Exceptions.ThrowGenericConversionNotSupported(
	sourceNamespaceName := NamespaceName,
	sourceClassName := ClassName,
	sourcePOUName := __POUNAME(),
	sourcePosition := __POSITION(),
	sourceDataType := TypeClass,
	targetDataType := otherValue.TypeClass
);
END_METHOD

(*!
<summary>Copies the stored byte representation into an equally sized target.</summary>
<description>
Requires a live writable target whose size equals Size. The caller is responsible for data compatibility: no
type check or numeric conversion is performed. Copies bytes from a nonzero Address referencing live source
storage. Does not clone referenced objects, transfer ownership, retain the target or modify this descriptor.
Copied pointer values still refer to the same resources and do not grant an independent right to release them.
A zero source Address raises DataMemberNotSpecifiedException without changing the target. A null target raises
ArgumentNotSpecifiedException; a target smaller than Size raises TargetVariableMemoryOverflowException; a
target larger than Size raises ArgumentOutOfRangeException before copying. Overlapping source and target
regions, including identical addresses, are supported through MEMMOVE. Descendants cannot override this
descriptor operation; customize value equality through IEqualityComparer or the stored object equality
contract.
</description>
*)
//!<param name="target">
//! Writable destination with the same byte size; its type interpretation is the caller's responsibility.
//! </param>
METHOD FINAL CopyTo
VAR_INPUT
	target : ANY;
END_VAR
IF Address = 0 THEN
	Exceptions.ThrowDataMemberNotSpecified(
		sourceNamespaceName := NamespaceName,
		sourceClassName := ClassName,
		sourcePOUName := __POUNAME(),
		sourcePosition := __POSITION(),
		dataMemberName := 'Address'
	);
END_IF

IF target.pValue = 0 THEN
	Exceptions.ThrowArgumentNotSpecified(
		sourceNamespaceName := NamespaceName,
		sourceClassName := ClassName,
		sourcePOUName := __POUNAME(),
		sourcePosition := __POSITION(),
		argumentName := 'target'
	); 
END_IF

IF TO_ULINT(target.diSize) < Size THEN
	Exceptions.ThrowTargetVariableMemoryOverflow(
		sourceNamespaceName := NamespaceName,
		sourceClassName := ClassName,
		sourcePOUName := __POUNAME(),
		sourcePosition := __POSITION(),
		targetVariableName := 'target.diSize',
		targetVariableSize := TO_ULINT(target.diSize)
	);
ELSIF TO_ULINT(target.diSize) > Size THEN
	Exceptions.ThrowArgumentOutOfRange(
		sourceNamespaceName := NamespaceName,
		sourceClassName := ClassName,
		sourcePOUName := __POUNAME(),
		sourcePosition := __POSITION(),
		argumentName := 'target.diSize',
		argumentValue := target.diSize
	);
END_IF

internalCopyTo(targetAddress := target.pValue);
END_METHOD

(*!
<summary>Compares generic values using an optional comparer or the built-in equality rules.</summary>
<description>
When comparer is supplied, AreEqual receives copies of both GENERIC_VALUE descriptors before any built-in
empty or type checks. OBJECT and USER_DEFINED remain distinct and Size is passed without conversion to
AnyType. The caller selects a compatible equality strategy, including its treatment of empty operands, and
keeps it and the data alive for the call. Comparer exceptions propagate without fallback. The comparer and
operands are borrowed only for the call; no payload is copied, cloned or released, and no ownership is
transferred. IsMemoryOwner does not affect the strategy's equality result. A supplied strategy must provide
GetValueHashCode consistent with AreEqual; this method does not compute a hash. Without a comparer, the
following built-in rules apply. INT_8 through INT_64 and UINT_8 through UINT_64 compare by value across widths
and signedness without floating-point conversion. A negative signed value never equals an unsigned value.
Pairs of REAL_32/REAL_64 values compare by canonical binary64 representation after widening non-NaN REAL
values, without a tolerance: positive and negative zero are equal, and all NaN encodings compare equal to each
other, including across widths, but not to non-NaN values. NaN is classified from integer bit views before
widening; other REAL widening follows the runtime floating-point configuration. A nonempty integer value and a
nonempty floating-point value always compare unequal, in either operand order. Both empty descriptors compare
equal; one empty descriptor compares unequal to a nonempty one. For nonempty descriptors, different TypeClass
values compare unequal except for the integer and floating-point pairs described above. BOOLEAN values compare
logically. Nonempty OBJECT descriptors delegate to the first live Object instance's Equals with the second
instance as its argument. The object type must provide a symmetric, transitive equality relation and a
matching GetHashCode; base Object uses identity equality. Callbacks and their exceptions propagate without
fallback. An address does not validate object lifetime. Other matching categories retain byte comparison:
strings use their actual string sizes, otherwise descriptor sizes are used. Dates and times compare by
representation only within the same TypeClass. Byte comparison covers the full ULINT length in bounded MEMCMP
chunks. USER_DEFINED compares all Size bytes, including padding and stored pointer values; equal fields do not
necessarily imply equal bytes, and the concrete user-defined type identity is not checked. Supply a compatible
comparer for field-based equality. Both descriptors must reference live storage consistent with their type and
size; no ownership is transferred. Descendants cannot override this descriptor operation; customize value
equality through IEqualityComparer or the stored object equality contract.
</description>
*)
//!<param name="otherValue">Descriptor of the value to compare.</param>
//!<param name="comparer">Optional borrowed equality and hashing strategy; zero selects built-in equality.</param>
METHOD FINAL Equals : BOOL
VAR_INPUT
	otherValue : GENERIC_VALUE;
	comparer : IEqualityComparer := 0;
END_VAR
VAR
	signedValue : LINT;

	firstObject : POINTER TO Object;
	secondObject : POINTER TO Object;

	stringPointer : POINTER TO STRING;
	wideStringPointer : POINTER TO WSTRING;
	referenceDataSize : ULINT;
	valueToCompareDataSize : ULINT;
	comparedSize : ULINT;
	chunkSize : UDINT;
END_VAR
IF comparer <> 0 THEN
	Equals := comparer.AreEqual(first := THIS^, second := otherValue);
	
	RETURN;
END_IF

IF IsNull OR_ELSE otherValue.IsNull THEN
	Equals := IsNull AND_THEN otherValue.IsNull;
ELSE
	CASE TypeClass OF
		GENERIC_TYPE_CLASS.INT_8, GENERIC_TYPE_CLASS.INT_16, GENERIC_TYPE_CLASS.INT_32, GENERIC_TYPE_CLASS.INT_64:
			CASE otherValue.TypeClass OF
				GENERIC_TYPE_CLASS.INT_8, GENERIC_TYPE_CLASS.INT_16, GENERIC_TYPE_CLASS.INT_32, GENERIC_TYPE_CLASS.INT_64:
					Equals := AsLInt() = otherValue.AsLInt();
					RETURN;

				GENERIC_TYPE_CLASS.UINT_8, GENERIC_TYPE_CLASS.UINT_16, GENERIC_TYPE_CLASS.UINT_32, GENERIC_TYPE_CLASS.UINT_64:
					signedValue := AsLInt();
					Equals := signedValue >= SignedInt64.ZERO AND_THEN TO_ULINT(signedValue) = otherValue.AsULInt();
					RETURN;
			END_CASE

		GENERIC_TYPE_CLASS.UINT_8, GENERIC_TYPE_CLASS.UINT_16, GENERIC_TYPE_CLASS.UINT_32, GENERIC_TYPE_CLASS.UINT_64:
			CASE otherValue.TypeClass OF
				GENERIC_TYPE_CLASS.INT_8, GENERIC_TYPE_CLASS.INT_16, GENERIC_TYPE_CLASS.INT_32, GENERIC_TYPE_CLASS.INT_64:
					signedValue := otherValue.AsLInt();
					Equals := signedValue >= SignedInt64.ZERO AND_THEN AsULInt() = TO_ULINT(signedValue);
					RETURN;

				GENERIC_TYPE_CLASS.UINT_8, GENERIC_TYPE_CLASS.UINT_16, GENERIC_TYPE_CLASS.UINT_32, GENERIC_TYPE_CLASS.UINT_64:
					Equals := AsULInt() = otherValue.AsULInt();
					RETURN;
			END_CASE

		GENERIC_TYPE_CLASS.REAL_32, GENERIC_TYPE_CLASS.REAL_64:
			CASE otherValue.TypeClass OF
				GENERIC_TYPE_CLASS.REAL_32, GENERIC_TYPE_CLASS.REAL_64:
					Equals := getCanonicalRealBits() = otherValue.getCanonicalRealBits();
					RETURN;
			END_CASE
	END_CASE

	IF TypeClass <> otherValue.TypeClass THEN
		Equals := FALSE;
		RETURN;
	END_IF

	IF TypeClass = GENERIC_TYPE_CLASS.OBJECT THEN
		firstObject := Address;
		secondObject := otherValue.Address;
		Equals := firstObject^.Equals(other := secondObject^);
		RETURN;
	END_IF

	IF TypeClass = GENERIC_TYPE_CLASS.BOOLEAN THEN
		Equals := AsBool() = otherValue.AsBool();
		RETURN;
	END_IF

	IF TypeClass = GENERIC_TYPE_CLASS.STRING_8 AND_THEN otherValue.TypeClass = GENERIC_TYPE_CLASS.STRING_8 THEN
		stringPointer := Address;
		referenceDataSize := Strings.GetActualSize(value := stringPointer^);
		
		stringPointer := otherValue.Address;		
		valueToCompareDataSize := Strings.GetActualSize(value := stringPointer^);
	ELSIF TypeClass = GENERIC_TYPE_CLASS.STRING_16 AND_THEN otherValue.TypeClass = GENERIC_TYPE_CLASS.STRING_16 THEN
		wideStringPointer := Address;
		referenceDataSize := WideStrings.GetActualSize(value := wideStringPointer^);
		
		wideStringPointer := otherValue.Address;		
		valueToCompareDataSize := WideStrings.GetActualSize(value := wideStringPointer^);
	ELSE
		referenceDataSize := Size;
		valueToCompareDataSize := otherValue.Size;		
	END_IF
 
	IF referenceDataSize <> valueToCompareDataSize THEN
		Equals := FALSE;
		RETURN;
	END_IF

	comparedSize := 0;

	WHILE comparedSize < referenceDataSize DO
		chunkSize := TO_UDINT(MIN(referenceDataSize - comparedSize, TO_ULINT(UnsignedInt32.MAX_VALUE)));

		IF Tc2_System.MEMCMP(
			pBuf1 := Address + TO_LWORD(comparedSize),
			pBuf2 := otherValue.Address + TO_LWORD(comparedSize),
			n := chunkSize
		) <> SignedInt32.ZERO THEN
			Equals := FALSE;
			RETURN;
		END_IF

		comparedSize := comparedSize + TO_ULINT(chunkSize);
	END_WHILE

	Equals := TRUE;
END_IF
END_METHOD

(*!
<summary>Returns a shared binary64 representation for generic floating-point equality and hashing.</summary>
<description>
Requires nonempty REAL_32 or REAL_64 storage of the matching representation. The typed Core operation classifies NaN from bits
before any floating conversion, maps all NaN encodings to one value, widens other REAL values to LREAL,
and maps both signed zeros to positive zero. Payload and ownership are unchanged. Widening follows the runtime
floating-point configuration.
</description>
*)
METHOD PRIVATE getCanonicalRealBits : ULINT
VAR
	valuePointer : UNIVERSAL_POINTER;
END_VAR
valuePointer.AsByte := Address;

IF TypeClass = GENERIC_TYPE_CLASS.REAL_32 THEN
	getCanonicalRealBits := Reals.GetCanonicalBinary64Bits(value := valuePointer.AsReal^);
ELSE
	getCanonicalRealBits := LongReals.GetCanonicalBinary64Bits(value := valuePointer.AsLReal^);
END_IF
END_METHOD

(*!
<summary>Computes a hash consistent with generic value equality or a supplied equality strategy.</summary>
<description>
A supplied comparer takes precedence even for empty descriptors; its GetValueHashCode exceptions propagate
without fallback. Use the same strategy for Equals and hashing. Without a comparer, empty descriptors hash to
zero. Integers are widened to 64-bit integer representations so equal values across widths and signedness hash
alike; negative signed integers are never equal to unsigned values. BOOLEAN is normalized to zero or one. REAL
values are widened to LREAL, both signed zeros are normalized, and all NaN encodings share one hash. Nonempty
OBJECT delegates to the live object's GetHashCode and requires its Equals/hash pair to agree. Strings hash
their actual terminated byte sequence, independent of storage capacity. Other categories hash all Size bytes,
matching the representation equality rules; USER_DEFINED includes padding and pointer fields and carries no
concrete type identity. The caller supplies live storage matching TypeClass and Size and keeps
equality-relevant data stable while a hash index uses it. IsMemoryOwner does not participate. Descriptors and
payload are borrowed without mutation, cloning, release or retained references. No instance fields, cached
hashes or dynamic allocations are introduced by the built-in hashing algorithm; user callbacks may have their
own costs and failures. The built-in byte hash uses FNV-1a with an explicitly masked 64-bit intermediate,
without relying on arithmetic overflow. Collisions are allowed and must be resolved with Equals. Hashes are
not persistent identifiers or portable serialization values. Runtime is proportional to the hashed byte count;
object and comparer callbacks define their own cost. Descendants cannot override this descriptor operation;
customize value equality through IEqualityComparer or the stored object equality contract.
</description>
*)
//!<param name="comparer">Optional borrowed equality and hashing strategy; zero selects the built-in rules.</param>
METHOD FINAL GetHashCode : UDINT
VAR_INPUT
	comparer : IEqualityComparer := 0;
END_VAR
VAR CONSTANT
	HASH_OFFSET_BASIS : UDINT := UDINT#2166136261;
	HASH_PRIME : ULINT := ULINT#16777619;
END_VAR
VAR
	signedValue : LINT;
	unsignedValue : ULINT;
	objectPointer : POINTER TO Object;
	stringPointer : POINTER TO STRING;
	wideStringPointer : POINTER TO WSTRING;

	dataPointer : POINTER TO BYTE;
	bytePointer : POINTER TO BYTE;
	dataSize : ULINT;
	index : ULINT;
	hashValue : UDINT;
	hashProduct : ULINT;
END_VAR
IF comparer <> 0 THEN
	GetHashCode := comparer.GetValueHashCode(value := THIS^);
	RETURN;
END_IF

IF IsNull THEN
	GetHashCode := 0;
	RETURN;
END_IF

dataPointer := Address;
dataSize := Size;

CASE TypeClass OF
	GENERIC_TYPE_CLASS.BOOLEAN:
		IF AsBool() THEN
			unsignedValue := 1;
		ELSE
			unsignedValue := 0;
		END_IF

		dataPointer := ADR(unsignedValue);
		dataSize := XSIZEOF(unsignedValue);

	GENERIC_TYPE_CLASS.INT_8, GENERIC_TYPE_CLASS.INT_16, GENERIC_TYPE_CLASS.INT_32, GENERIC_TYPE_CLASS.INT_64:
		signedValue := AsLInt();
		dataPointer := ADR(signedValue);
		dataSize := XSIZEOF(signedValue);

	GENERIC_TYPE_CLASS.UINT_8, GENERIC_TYPE_CLASS.UINT_16, GENERIC_TYPE_CLASS.UINT_32, GENERIC_TYPE_CLASS.UINT_64:
		unsignedValue := AsULInt();
		dataPointer := ADR(unsignedValue);
		dataSize := XSIZEOF(unsignedValue);

	GENERIC_TYPE_CLASS.REAL_32, GENERIC_TYPE_CLASS.REAL_64:
		unsignedValue := getCanonicalRealBits();
		dataPointer := ADR(unsignedValue);
		dataSize := XSIZEOF(unsignedValue);

	GENERIC_TYPE_CLASS.STRING_8:
		stringPointer := Address;
		dataSize := Strings.GetActualSize(value := stringPointer^);

	GENERIC_TYPE_CLASS.STRING_16:
		wideStringPointer := Address;
		dataSize := WideStrings.GetActualSize(value := wideStringPointer^);

	GENERIC_TYPE_CLASS.OBJECT:
		objectPointer := Address;
		GetHashCode := objectPointer^.GetHashCode();
		RETURN;
END_CASE

hashValue := HASH_OFFSET_BASIS;
index := 0;

WHILE index < dataSize DO
	bytePointer := dataPointer + TO_LWORD(index);
	hashProduct := TO_ULINT(hashValue XOR TO_UDINT(bytePointer^)) * HASH_PRIME;
	hashValue := TO_UDINT(hashProduct AND TO_ULINT(UnsignedInt32.MAX_VALUE));
	index := index + 1;
END_WHILE

GetHashCode := hashValue;
END_METHOD

(*!
<summary>Copies the payload bytes to a destination already checked by the caller.</summary>
<description>
The destination must be writable for Size bytes. Address must be nonzero and reference readable storage of
that size; overlapping regions are supported. The caller checks for a zero source address before calling. No
cloning or ownership transfer is performed.
</description>
*)
METHOD PRIVATE internalCopyTo
VAR_INPUT
	targetAddress : PVOID;
END_VAR
Tc2_System.MEMMOVE(destAddr := targetAddress, srcAddr := Address, n := TO_UDINT(Size));
END_METHOD

(*!
<summary>Checks whether an As* accessor supports the source and target representation pair.</summary>
<description>
Inspects TypeClass only, without reading payload storage, allocating memory or raising exceptions. TRUE means
that a matching conversion branch exists; it does not guarantee a live value, sufficient storage, an in-range
result or lossless conversion. The selected As* accessor still applies its value checks and loss flag. Returns
FALSE for unsupported pairs, including OBJECT to text and targets without an As* accessor. No conversion is
performed and no ownership is transferred.
</description>
*)
//!<param name="targetTypeClass">Desired target generic representation category.</param>
METHOD FINAL IsConvertibleTo : BOOL
VAR_INPUT
	targetTypeClass : GENERIC_TYPE_CLASS;
END_VAR
CASE targetTypeClass OF
	GENERIC_TYPE_CLASS.BOOLEAN,
	GENERIC_TYPE_CLASS.INT_16,
	GENERIC_TYPE_CLASS.INT_32,
	GENERIC_TYPE_CLASS.INT_64,
	GENERIC_TYPE_CLASS.UINT_8,
	GENERIC_TYPE_CLASS.UINT_16,
	GENERIC_TYPE_CLASS.UINT_32,
	GENERIC_TYPE_CLASS.UINT_64:
		IsConvertibleTo := TypeClass >= GENERIC_TYPE_CLASS.BOOLEAN AND_THEN TypeClass <= GENERIC_TYPE_CLASS.UINT_64;

	GENERIC_TYPE_CLASS.INT_8:
		IsConvertibleTo := (TypeClass >= GENERIC_TYPE_CLASS.INT_8 AND_THEN TypeClass <= GENERIC_TYPE_CLASS.INT_64)
			OR_ELSE (TypeClass >= GENERIC_TYPE_CLASS.UINT_16 AND_THEN TypeClass <= GENERIC_TYPE_CLASS.UINT_64);

	GENERIC_TYPE_CLASS.REAL_32:
		IsConvertibleTo := TypeClass = GENERIC_TYPE_CLASS.REAL_32 OR_ELSE TypeClass = GENERIC_TYPE_CLASS.REAL_64;

	GENERIC_TYPE_CLASS.REAL_64:
		IsConvertibleTo := TypeClass >= GENERIC_TYPE_CLASS.BOOLEAN AND_THEN TypeClass <= GENERIC_TYPE_CLASS.REAL_64;

	GENERIC_TYPE_CLASS.STRING_8,
	GENERIC_TYPE_CLASS.STRING_16:
		IsConvertibleTo := TypeClass >= GENERIC_TYPE_CLASS.BOOLEAN AND_THEN TypeClass <= GENERIC_TYPE_CLASS.TIME_OF_DAY_64;

	GENERIC_TYPE_CLASS.DATE_32:
		IsConvertibleTo := TypeClass = GENERIC_TYPE_CLASS.DATE_32
			OR_ELSE TypeClass = GENERIC_TYPE_CLASS.DATE_64
			OR_ELSE TypeClass = GENERIC_TYPE_CLASS.DATE_AND_TIME_32
			OR_ELSE TypeClass = GENERIC_TYPE_CLASS.INT_32
			OR_ELSE TypeClass = GENERIC_TYPE_CLASS.UINT_32
			OR_ELSE TypeClass = GENERIC_TYPE_CLASS.INT_64
			OR_ELSE TypeClass = GENERIC_TYPE_CLASS.UINT_64;

	GENERIC_TYPE_CLASS.DATE_64:
		IsConvertibleTo := TypeClass = GENERIC_TYPE_CLASS.DATE_32
			OR_ELSE TypeClass = GENERIC_TYPE_CLASS.DATE_64
			OR_ELSE TypeClass = GENERIC_TYPE_CLASS.DATE_AND_TIME_32
			OR_ELSE TypeClass = GENERIC_TYPE_CLASS.DATE_AND_TIME_64
			OR_ELSE TypeClass = GENERIC_TYPE_CLASS.INT_64
			OR_ELSE TypeClass = GENERIC_TYPE_CLASS.UINT_64;

	GENERIC_TYPE_CLASS.DATE_AND_TIME_32:
		IsConvertibleTo := TypeClass = GENERIC_TYPE_CLASS.DATE_32
			OR_ELSE TypeClass = GENERIC_TYPE_CLASS.DATE_AND_TIME_32
			OR_ELSE TypeClass = GENERIC_TYPE_CLASS.DATE_AND_TIME_64
			OR_ELSE TypeClass = GENERIC_TYPE_CLASS.INT_32
			OR_ELSE TypeClass = GENERIC_TYPE_CLASS.UINT_32
			OR_ELSE TypeClass = GENERIC_TYPE_CLASS.INT_64
			OR_ELSE TypeClass = GENERIC_TYPE_CLASS.UINT_64;

	GENERIC_TYPE_CLASS.DATE_AND_TIME_64:
		IsConvertibleTo := TypeClass = GENERIC_TYPE_CLASS.DATE_32
			OR_ELSE TypeClass = GENERIC_TYPE_CLASS.DATE_64
			OR_ELSE TypeClass = GENERIC_TYPE_CLASS.DATE_AND_TIME_32
			OR_ELSE TypeClass = GENERIC_TYPE_CLASS.DATE_AND_TIME_64
			OR_ELSE TypeClass = GENERIC_TYPE_CLASS.TIME_32
			OR_ELSE TypeClass = GENERIC_TYPE_CLASS.TIME_64
			OR_ELSE TypeClass = GENERIC_TYPE_CLASS.INT_64
			OR_ELSE TypeClass = GENERIC_TYPE_CLASS.UINT_64;

	GENERIC_TYPE_CLASS.TIME_32:
		IsConvertibleTo := TypeClass = GENERIC_TYPE_CLASS.TIME_32
			OR_ELSE TypeClass = GENERIC_TYPE_CLASS.TIME_64
			OR_ELSE TypeClass = GENERIC_TYPE_CLASS.TIME_OF_DAY_32
			OR_ELSE TypeClass = GENERIC_TYPE_CLASS.DATE_AND_TIME_32
			OR_ELSE TypeClass = GENERIC_TYPE_CLASS.INT_32
			OR_ELSE TypeClass = GENERIC_TYPE_CLASS.UINT_32
			OR_ELSE TypeClass = GENERIC_TYPE_CLASS.INT_64
			OR_ELSE TypeClass = GENERIC_TYPE_CLASS.UINT_64;

	GENERIC_TYPE_CLASS.TIME_64:
		IsConvertibleTo := TypeClass = GENERIC_TYPE_CLASS.TIME_32
			OR_ELSE TypeClass = GENERIC_TYPE_CLASS.TIME_64
			OR_ELSE TypeClass = GENERIC_TYPE_CLASS.TIME_OF_DAY_32
			OR_ELSE TypeClass = GENERIC_TYPE_CLASS.TIME_OF_DAY_64
			OR_ELSE TypeClass = GENERIC_TYPE_CLASS.DATE_AND_TIME_32
			OR_ELSE TypeClass = GENERIC_TYPE_CLASS.DATE_AND_TIME_64
			OR_ELSE TypeClass = GENERIC_TYPE_CLASS.INT_64
			OR_ELSE TypeClass = GENERIC_TYPE_CLASS.UINT_64;

	GENERIC_TYPE_CLASS.TIME_OF_DAY_32:
		IsConvertibleTo := TypeClass = GENERIC_TYPE_CLASS.TIME_OF_DAY_32
			OR_ELSE TypeClass = GENERIC_TYPE_CLASS.TIME_32
			OR_ELSE TypeClass = GENERIC_TYPE_CLASS.TIME_64
			OR_ELSE TypeClass = GENERIC_TYPE_CLASS.INT_32
			OR_ELSE TypeClass = GENERIC_TYPE_CLASS.UINT_32
			OR_ELSE TypeClass = GENERIC_TYPE_CLASS.INT_64
			OR_ELSE TypeClass = GENERIC_TYPE_CLASS.UINT_64;

	GENERIC_TYPE_CLASS.TIME_OF_DAY_64:
		IsConvertibleTo := TypeClass = GENERIC_TYPE_CLASS.TIME_OF_DAY_32
			OR_ELSE TypeClass = GENERIC_TYPE_CLASS.TIME_OF_DAY_64
			OR_ELSE TypeClass = GENERIC_TYPE_CLASS.TIME_32
			OR_ELSE TypeClass = GENERIC_TYPE_CLASS.TIME_64
			OR_ELSE TypeClass = GENERIC_TYPE_CLASS.DATE_AND_TIME_32
			OR_ELSE TypeClass = GENERIC_TYPE_CLASS.DATE_AND_TIME_64
			OR_ELSE TypeClass = GENERIC_TYPE_CLASS.INT_64
			OR_ELSE TypeClass = GENERIC_TYPE_CLASS.UINT_64;

	GENERIC_TYPE_CLASS.OBJECT:
		IsConvertibleTo := TypeClass = GENERIC_TYPE_CLASS.OBJECT;
END_CASE
END_METHOD

(*!
<summary>Reports whether the descriptor has no usable value metadata.</summary>
<description>
TRUE when TypeClass is UNSPECIFIED, Address is zero or Size is zero. This is the empty-value criterion used by
built-in Equals and GetHashCode; a supplied comparer defines its own policy. It does not validate payload
lifetime or address validity. An empty descriptor may still own allocated storage; IsNull does not remove the
obligation to Release it.
</description>
*)
{attribute 'monitoring' := 'call'}
PROPERTY FINAL IsNull : BOOL
GET
IsNull := TypeClass = GENERIC_TYPE_CLASS.UNSPECIFIED OR_ELSE Address = 0 OR_ELSE Size = 0;
END_GET
END_PROPERTY

(*!
<summary>Provides the library namespace used in diagnostics.</summary>
<description>
Borrowed read-only reference to the compiler-initialized library namespace; no ownership transfer.
</description>
*)
{attribute 'monitoring' := 'call'}
PROPERTY NamespaceName : REFERENCE TO STRING
GET
NamespaceName REF= CurrentNamespace.Name;
END_GET
END_PROPERTY

(*!
<summary>Attempts release of owned storage and resets the descriptor.</summary>
<description>
Borrowed storage is not freed. Owned objects use the object-release path; other owned storage uses raw-memory
release. The descriptor is reset even if TryReleaseDynamicMemory fails; successful deallocation is not
guaranteed and other aliases are not cleared. Descendants cannot override this descriptor operation; customize
value equality through IEqualityComparer or the stored object equality contract.
</description>
*)
METHOD FINAL Release
IF IsMemoryOwner THEN
	Memory.TryReleaseDynamicMemory(address := Address, isObject := TypeClass = GENERIC_TYPE_CLASS.OBJECT);
END_IF

Reset();
END_METHOD

(*!
<summary>Clears type, address, size and ownership metadata without freeing memory.</summary>
<description>
Use after transferring ownership or when no owned storage remains. Resetting an owning descriptor without
arranging release loses its ownership information; no destructor or allocation is performed. Descendants
cannot override this descriptor operation; customize value equality through IEqualityComparer or the stored
object equality contract.
</description>
*)
METHOD FINAL Reset
TypeClass := GENERIC_TYPE_CLASS.UNSPECIFIED;
Address := 0;
Size := 0;
IsMemoryOwner := FALSE;
END_METHOD

(*!
<summary>Attempts to copy a compatible value into the existing generic storage.</summary>
<description>
Unsupported types, incompatible storage and copy failure return FALSE without creating a diagnostic exception.
Native exceptions are contained. A latched allocation failure returns FALSE.
Does not change descriptor fields or transfer ownership.
Requires live source and destination storage; copied bytes are not rolled back on failure. Preserves terminal
allocation state for the task boundary. Descendants cannot override this descriptor operation; customize value
equality through IEqualityComparer or the stored object equality contract.
</description>
*)
METHOD FINAL TryChangeValueByAny : BOOL
VAR_INPUT
	value : ANY;
	isObject : BOOL := FALSE;
END_VAR
TryChangeValueByAny := TryChangeValueByAnyType(value := value, isObject := isObject);
END_METHOD

(*!
<summary>Attempts to copy a compatible value into the existing generic storage.</summary>
<description>
Unsupported types, incompatible storage and copy failure return FALSE without creating a diagnostic exception.
Native exceptions are contained. A latched allocation failure returns FALSE.
Does not change descriptor fields or transfer ownership.
Requires live source and destination storage; copied bytes are not rolled back on failure. Preserves terminal
allocation state for the task boundary. Descendants cannot override this descriptor operation; customize value
equality through IEqualityComparer or the stored object equality contract.
</description>
*)
METHOD FINAL TryChangeValueByAnyType : BOOL
VAR_INPUT
	value : __SYSTEM.AnyType;
	isObject : BOOL := FALSE;
END_VAR
VAR
	sourceType : GENERIC_TYPE_CLASS;
END_VAR
IF DynamicMemoryManager.HasAllocationFailed THEN
	RETURN;
END_IF

__TRY
	IF GenericTypeClassConvertor.TryGetGenericTypeClassBySystemAnyType(
		systemAnyType := value,
		isObject := isObject,
		genericTypeClass => sourceType
	)
	THEN
		TryChangeValueByAnyType := copyMappedValue(value := value, sourceType := sourceType)
			= GENERIC_VALUE_COPY_RESULT.COPIED;
	END_IF
__CATCH
	TryChangeValueByAnyType := FALSE;
__ENDTRY

IF DynamicMemoryManager.HasAllocationFailed THEN
	TryChangeValueByAnyType := FALSE;
END_IF
END_METHOD

(*!
<summary>Copies the byte representation when the target address and size are acceptable.</summary>
<description>
Returns FALSE without copying for a zero source Address, a null target or a size mismatch; otherwise copies
and returns TRUE. The caller supplies live writable storage and is responsible for data compatibility. No type
conversion, cloning or ownership transfer is performed. Overlapping regions, including identical addresses,
are supported. Catches exceptions and returns FALSE. A failed memory operation can leave partially copied
bytes; no rollback is performed. Catching an exception does not validate memory lifetime. Descendants cannot
override this descriptor operation; customize value equality through IEqualityComparer or the stored object
equality contract.
</description>
*)
//!<param name="target">Writable destination with the same byte size.</param>
METHOD FINAL TryCopyTo : BOOL
VAR_INPUT
	target : ANY;
END_VAR
__TRY
	IF Address = 0 OR_ELSE target.pValue = 0 THEN
		RETURN; 
	END_IF

	IF TO_ULINT(target.diSize) <> Size THEN
		RETURN; 
	END_IF

	internalCopyTo(targetAddress := target.pValue);

	TryCopyTo := TRUE;
__CATCH
	TryCopyTo := FALSE;
__ENDTRY
END_METHOD

END_FUNCTION_BLOCK

(* stored: Version 1.1.0.1
   POU GENERIC_VALUE: Id {4ec776d3-51b8-42d3-97bb-5e4d1a102b1f}, SpecialFunc None
   Folder AsTyped: Id {e96a41ac-e3cd-4eee-9bfa-b62dba0c2d0e}
   Folder Date and time: Id {0e8135f9-c7a8-41d0-996d-4e135d2a2366}
   Folder Floating point: Id {8039a744-40ce-4546-beea-78a288e45706}
   Folder Integer: Id {e3759741-5c8c-482f-93b9-6ae90a2f6296}
   Folder Signed: Id {fb335c0b-7655-449f-bc46-48fb10ad905c}
   Folder Unsugned: Id {bab4b970-dedd-4b75-8710-280ec540561b}
   Folder Strings: Id {f6373c83-d47f-4dab-9f39-83ae4e8a3796}
   Folder ChangeValue: Id {ff6ec9ec-7e82-4906-a7b3-4f1a0bbc2daf}
   Folder CleanupMethods: Id {6633f1de-b2f9-411c-a1ba-5eaade50e25e}
   Folder Service methods: Id {f60d642b-cec1-4cae-991f-d82121762e9d}
   Method AsAnyType: Id {59db7a53-29a2-4c5e-a06f-b2b343ab8f25}
   Method AsBool: Id {1aaa60f7-a8aa-48fc-a4c3-f53925263a40}
   Method AsByte: Id {936f9e9f-e35c-461b-a5b6-c2e02b118baf}
   Method AsDate: Id {db320a05-493c-45cf-92f8-51bf496ee511}
   Method AsDateAndTime: Id {ba931761-c96e-42e2-9fa4-d1882172beda}
   Method AsDInt: Id {4fea0b7d-fe5e-4808-9a02-b0a72b1114c9}
   Method AsDWord: Id {1ee84003-88d5-466d-8c56-9b5d650c16eb}
   Method AsInt: Id {fbd81b42-6af9-470c-9770-5641903fbac8}
   Method AsIObject: Id {80096a9d-d283-480b-80a4-d0dd536beae0}
   Method AsLDate: Id {a43023c1-e686-4d4d-82c6-573f5b54a6de}
   Method AsLDateAndTime: Id {36a42bba-09cd-44d2-9d6f-f83ecf955631}
   Method AsLInt: Id {557ab87e-2262-4a71-b53a-324d552cca35}
   Method AsLReal: Id {6ff6d2d4-05a2-4a88-8dfa-3efa48fa159c}
   Method AsLTime: Id {312f2003-0852-4cfd-8313-e6043e172de5}
   Method AsLTimeOfDay: Id {3746ef26-79d9-476c-ba8d-9d1fb97744ec}
   Method AsLWord: Id {329d366e-53cb-444a-baae-0e3cbf144975}
   Method AsObject: Id {996e8fad-fcc2-4f05-b582-9a439f872e26}
   Method AsReal: Id {45160cf2-6e60-4035-806b-879e84f1bb89}
   Method Assign: Id {862ebf60-dfb4-45d8-a755-cbc5dc31a2cb}
   Method AsSInt: Id {17b44680-9119-41da-9958-f566e80539b5}
   Method AsString255: Id {34520551-01e7-4ae7-9a34-54ba8a2cf3c1}
   Method AsStringReference: Id {5ecee28b-da1c-4264-92ee-6c69f4328ec9}
   Method AsTime: Id {b0c8a8a8-d7c2-483f-b215-128f7d04ba16}
   Method AsTimeOfDay: Id {83f725a7-471b-4136-801c-36fbe6098098}
   Method AsUDInt: Id {90863b55-b5cf-4472-b2f4-3d7e5196f54f}
   Method AsUInt: Id {0cb7d9b1-a26c-4d44-8107-5807eda8eaa5}
   Method AsULInt: Id {ddfdd7f6-ff0f-4202-a7b9-d1b08069f76c}
   Method AsUSInt: Id {7f2825bd-7342-487e-96ac-27ff3bcc2e3c}
   Method AsWord: Id {5e995462-8574-4174-bafd-d9d8e8e626c5}
   Method AsWString255: Id {02ab723a-3f42-4d36-a0f6-c0e9871bfd09}
   Method AsWStringReference: Id {31493745-1b4b-4427-a5e6-18639dd644fb}
   Method ChangeValueByAny: Id {f7c7dd69-068a-47f7-bb61-709a535f4d37}
   Method copyMappedValue: Id {1314e191-897c-4c5d-8cd0-6938238073f2}
   Method ChangeValueByAnyType: Id {1e16a561-f4aa-4df6-80a7-92686d04f493}
   Property ClassName: Id {a1f78ed3-d25a-4e81-8b88-934a58828338}
   Get Get: Id {9652d94e-8909-435e-98b2-6d0f00f73d32}
   Method compareIntegerToReal: Id {219a7d64-fe46-45ab-9db1-f7c748e9fe60}
   Method CompareTo: Id {5ce2e755-e8a0-495e-b60d-5197776627f3}
   Method CopyTo: Id {a9e28a3d-762a-4fcd-99e6-4d377c8be6f0}
   Method Equals: Id {165ded56-3861-403f-9838-406d75321178}
   Method getCanonicalRealBits: Id {c0c43419-5c5f-48f3-bb40-f8d8b2204104}
   Method GetHashCode: Id {091c42af-fc6a-4c30-a170-e310c535bc0a}
   Method internalCopyTo: Id {dffcbd59-ee39-4c74-bc12-2c951ca57eee}
   Method IsConvertibleTo: Id {3876d0ba-dd7a-4ef3-bc6f-7b8542042d4e}
   Property IsNull: Id {b0a5dbd8-6fb5-436e-9b63-9e18aded8437}
   Get Get: Id {293dd0e0-6dfe-4234-9575-a1a778286228}
   Property NamespaceName: Id {6b1b9ffb-991c-4d04-a51f-7608d3745ab0}
   Get Get: Id {70ea020b-d8b3-4815-b692-efc03598f31f}
   Method Release: Id {9937fc92-8120-434b-ac91-5b20bd6f7de6}
   Method Reset: Id {7b456980-e70d-4684-918f-f6fc89768f34}
   Method TryChangeValueByAny: Id {27b8e08e-2fa6-41be-af60-419256c2188b}
   Method TryChangeValueByAnyType: Id {4ed65d07-87f2-4259-80eb-13281b15e53c}
   Method TryCopyTo: Id {ce4998f1-fc8d-443b-ab31-7fcdb66ae168} *)
